(* Logix 5000 project; controller R400_500_XLS vendor 1 type 14 code 216 rev 31.11; software revision 31.01; part 5 of 32 *)
(* tags used below, declared in another part *)
   Abort1 : DINT;   // Not Used
   Cycles : UDT_CYCLE[11];
   CycleSequence : UDT_CYCLE_SEQUENCE;
   I_Pw_Tnk_Lvl_Sw_Deb : BOOL;   // Debounced pure water tank level switch (100ms)
   M : DINT[5];   // Memory Bits
   MinorFaultCheck : TIMER;
   MinorFaultRecord : FaultRecord;
   OneShot : DINT[1];
   ONS_FC01 : DINT;
   ONS_FC11 : DINT;
   ONS_FC12 : DINT;
   ONS_FC13 : DINT;
   ONS_FC64 : DINT;
   ONS_WSH30 : SINT;
   ONS_WSH35 : SINT;
   Service : DINT[2];   // Unused Service Mode Memory Bit
   String : STRING[50];   // String
   Tmr : TIMER[107];
   Unld_Door : DINT;
   BatteryLowWarning : BOOL;
   bFactoryResetCompleted : BOOL;
   bONSSerialModuleResetInhibit : BOOL;
   bONSSerialModuleSetInhibit : BOOL;
   bSerialModuleConfigureInhibit : BOOL;   // Configure if Serial Card is Inhibited or not
   Cfg_10_Modules : BOOL;   // Chassis is configured 10 slots
   Cfg_11_Modules : BOOL;
   Chassis_Size_Ret : DINT[3];
   Ctrlr_Status : DINT;
   Current_Screen : DINT;
   DateTime : DINT[7];
   DISABLE : BOOL;   // Disable bit
   EmailSMSInt : INT[8];   // Email & SMS Notification Integer
   EnDis_LabWasher : DINT;
   EnDis_LabWasher2 : DINT;
   Ethernet_Config_Msg : MESSAGE;
   F8 : REAL[6];
   I_Chem_Cond : DINT;   // Chemical water conductivity
   I_Chm_1_Lvl_Sw : BOOL;   // Chemical Pump #1 level switch
   I_Chm_2_Lvl_Sw : BOOL;   // Chemical Pump #2 level switch
   I_Chm_3_Lvl_Sw : BOOL;   // Chemical Pump #3 level switch
   I_Chm_4_Lvl_Sw : BOOL;   // Chemical Pump #4 level switch
   I_Dry_RTD : DINT;   // Drying RTD
   I_Final_Rinse_Cond : DINT;   // Final rinse water conductivity
   I_Ld_Dr_Cls_Sw : BOOL;   // Load door close
   I_Ld_Dr_Obs_Sw : BOOL;   // Load door obstruction switch
   I_MCR : BOOL;   // MCR input
   I_Mtr_Ovrld : BOOL;   // Motor overload
   I_Pump_Press : DINT;   // Recirculation pump pressure
   I_Pure_Water_Filling_Auth : BOOL;
   I_Pw_Tnk_Lvl_Sw : BOOL;   // Pure water tank level switch
   I_Pw_Tnk_RTD : DINT;   // Pure water tank RTD
   I_Pw_Tnk_Sft_Lvl_Sw : BOOL;   // Pure water tank safety level switch
   I_Shlf_Sw : BOOL;   // Shelf switch
   I_Smp_Lvl_Hgh : BOOL;   // Sump high level switch
   I_Smp_Lvl_Lw : BOOL;   // Sump low level switch
   I_Smp_RTD : DINT;   // Sump RTD
   I_Smp_Sft_Lvl_Sw : BOOL;   // Sump safety level switch
   I_Unld_Dr_Cls_Sw : BOOL;   // Unload door close
   I_Unld_Dr_Obs_Sw : BOOL;   // Unload door obstruction switch
   I_UnldDr_ClseSlnce_Bttn : BOOL;   // Door Close/ Silence button Unload Side
   I_UnldDr_Opn_Bttn : BOOL;   // Door Open button Unload side
   iSerialModuleActivateDeactivateInhibit : DINT;   // Set Bit 2 Of Word to Inhibited Serial M Reset Bit 2 Of Word to Un-inhibited
   L32E_ETH_Cfg : TIMER;   // Delay for Ethernet port initialization
   Language_English : STRING;
   MinorFaultBits : DINT;
   msg : BOOL[512];
   Msg_PwrUp : DINT;
   N13 : DINT;
   NOT_USED : SINT[3];
   ONS_WSH64 : SINT;
   previous_s108 : DINT;
   RD_CHASSIS_1 : MESSAGE;
   RD_CHASSIS_2 : MESSAGE;
   RemoteDisplayNumber : DINT;   // HMI connection
   sChangeLanguage : STRING;   // jplv09
   Screen_Ctrl : DINT;   // PLC Screen Request
   SimGenEnabled : BOOL;   // SimGen enable bit 1= Simgen ON
   Tpb : DINT[11];
   TpbImage : DINT[11];
   Unit : Hrdwre;   // Unit Configuration
   WR_CHASSIS_10 : MESSAGE;
   WR_CHASSIS_11 : MESSAGE;
(* MainProgram, continued *)

ROUTINE Inputs_10_Modules   (* ladder *)
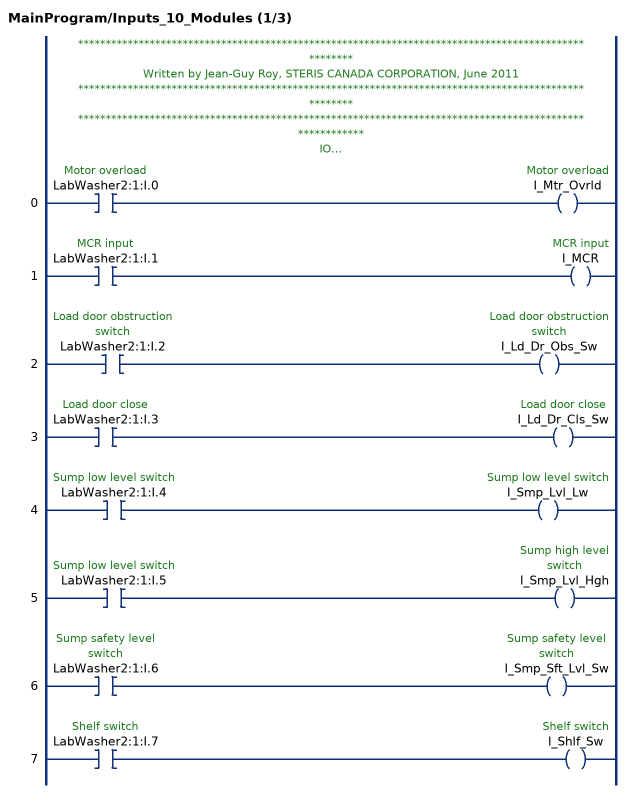
   // ****************************************************************************************************
   // Written by Jean-Guy Roy, STERIS CANADA CORPORATION, June 2011
   // ****************************************************************************************************
   // ********************************************************************************************************
   // IO1
   // ********************************************************************************************************
   0: XIC(LabWasher2:1:I.0)OTE(I_Mtr_Ovrld);
   1: XIC(LabWasher2:1:I.1)OTE(I_MCR);
   2: XIC(LabWasher2:1:I.2)OTE(I_Ld_Dr_Obs_Sw);
   3: XIC(LabWasher2:1:I.3)OTE(I_Ld_Dr_Cls_Sw);
   4: XIC(LabWasher2:1:I.4)OTE(I_Smp_Lvl_Lw);
   5: XIC(LabWasher2:1:I.5)OTE(I_Smp_Lvl_Hgh);
   6: XIC(LabWasher2:1:I.6)OTE(I_Smp_Sft_Lvl_Sw);
   7: XIC(LabWasher2:1:I.7)OTE(I_Shlf_Sw);
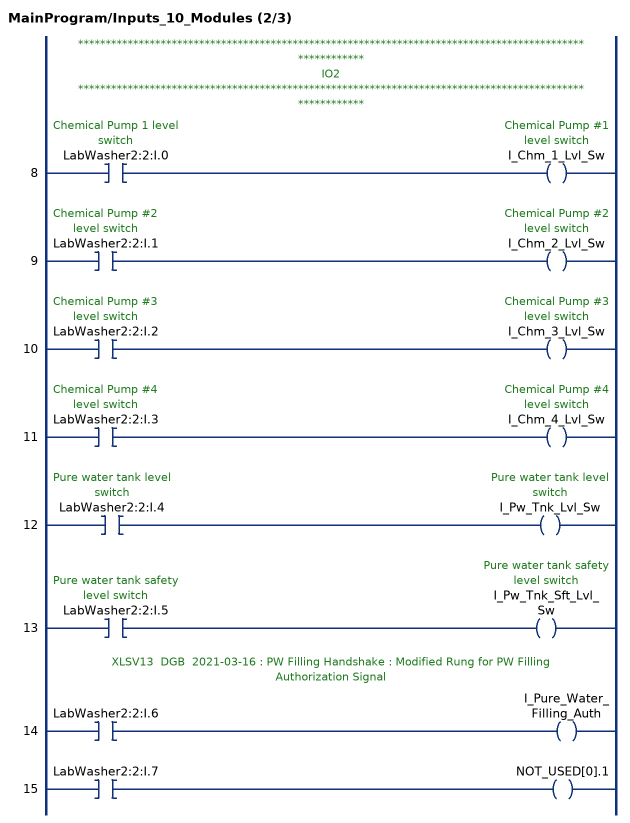
   // ********************************************************************************************************
   // IO2
   // ********************************************************************************************************
   8: XIC(LabWasher2:2:I.0)OTE(I_Chm_1_Lvl_Sw);
   9: XIC(LabWasher2:2:I.1)OTE(I_Chm_2_Lvl_Sw);
   10: XIC(LabWasher2:2:I.2)OTE(I_Chm_3_Lvl_Sw);
   11: XIC(LabWasher2:2:I.3)OTE(I_Chm_4_Lvl_Sw);
   12: XIC(LabWasher2:2:I.4)OTE(I_Pw_Tnk_Lvl_Sw);
   13: XIC(LabWasher2:2:I.5)OTE(I_Pw_Tnk_Sft_Lvl_Sw);
   // XLSV13  DGB  2021-03-16 : PW Filling Handshake : Modified Rung for PW Filling Authorization Signal
   14: XIC(LabWasher2:2:I.6)OTE(I_Pure_Water_Filling_Auth);
   15: XIC(LabWasher2:2:I.7)OTE(NOT_USED[0].1);
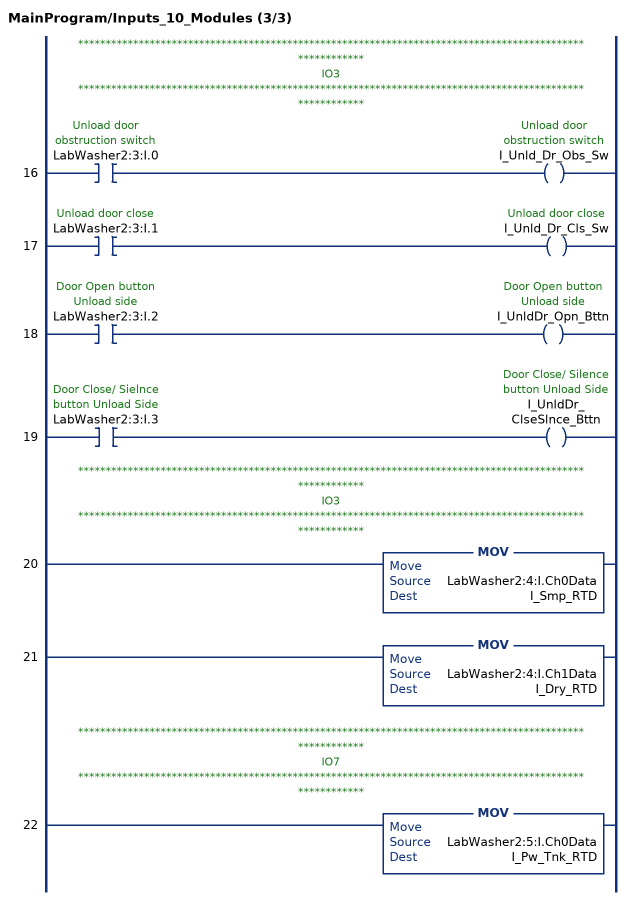
   // ********************************************************************************************************
   // IO3
   // ********************************************************************************************************
   16: XIC(LabWasher2:3:I.0)OTE(I_Unld_Dr_Obs_Sw);
   17: XIC(LabWasher2:3:I.1)OTE(I_Unld_Dr_Cls_Sw);
   18: XIC(LabWasher2:3:I.2)OTE(I_UnldDr_Opn_Bttn);
   19: XIC(LabWasher2:3:I.3)OTE(I_UnldDr_ClseSlnce_Bttn);
   // ********************************************************************************************************
   // IO3
   // ********************************************************************************************************
   20: MOV(LabWasher2:4:I.Ch0Data,I_Smp_RTD);
   21: MOV(LabWasher2:4:I.Ch1Data,I_Dry_RTD);
   // ********************************************************************************************************
   // IO7
   // ********************************************************************************************************
   22: MOV(LabWasher2:5:I.Ch0Data,I_Pw_Tnk_RTD);
END_ROUTINE

ROUTINE Inputs_Debounced   (* ladder *)
// This routine manages the debounced inputs
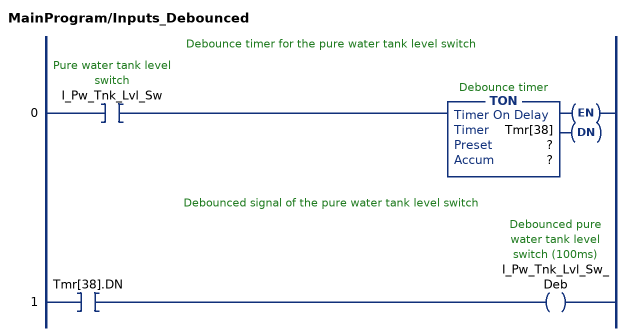
   // Debounce timer for the pure water tank level switch
   0: XIC(I_Pw_Tnk_Lvl_Sw)TON(Tmr[38],?,?);
   // Debounced signal of the pure water tank level switch
   1: XIC(Tmr[38].DN)OTE(I_Pw_Tnk_Lvl_Sw_Deb);
END_ROUTINE

ROUTINE Inputs_Smgn   (* ladder *)
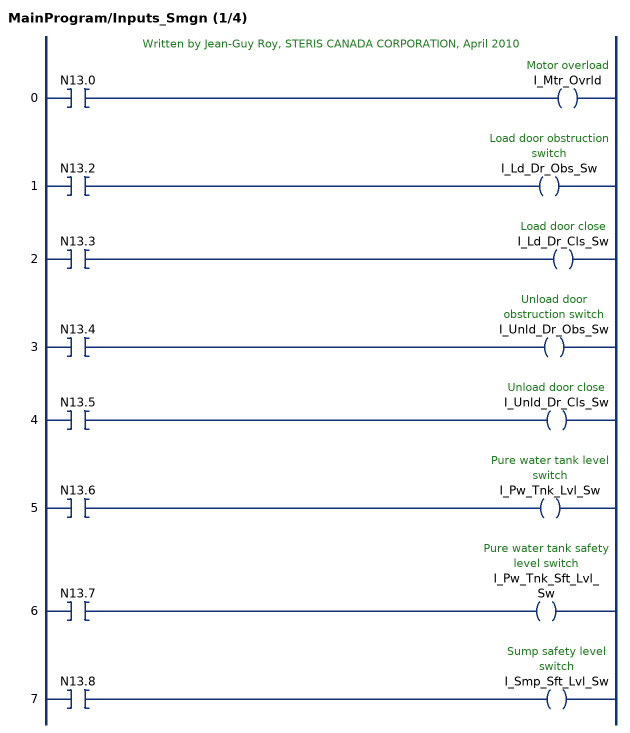
   // Written by Jean-Guy Roy, STERIS CANADA CORPORATION, April 2010
   0: XIC(N13.0)OTE(I_Mtr_Ovrld);
   1: XIC(N13.2)OTE(I_Ld_Dr_Obs_Sw);
   2: XIC(N13.3)OTE(I_Ld_Dr_Cls_Sw);
   3: XIC(N13.4)OTE(I_Unld_Dr_Obs_Sw);
   4: XIC(N13.5)OTE(I_Unld_Dr_Cls_Sw);
   5: XIC(N13.6)OTE(I_Pw_Tnk_Lvl_Sw);
   6: XIC(N13.7)OTE(I_Pw_Tnk_Sft_Lvl_Sw);
   7: XIC(N13.8)OTE(I_Smp_Sft_Lvl_Sw);
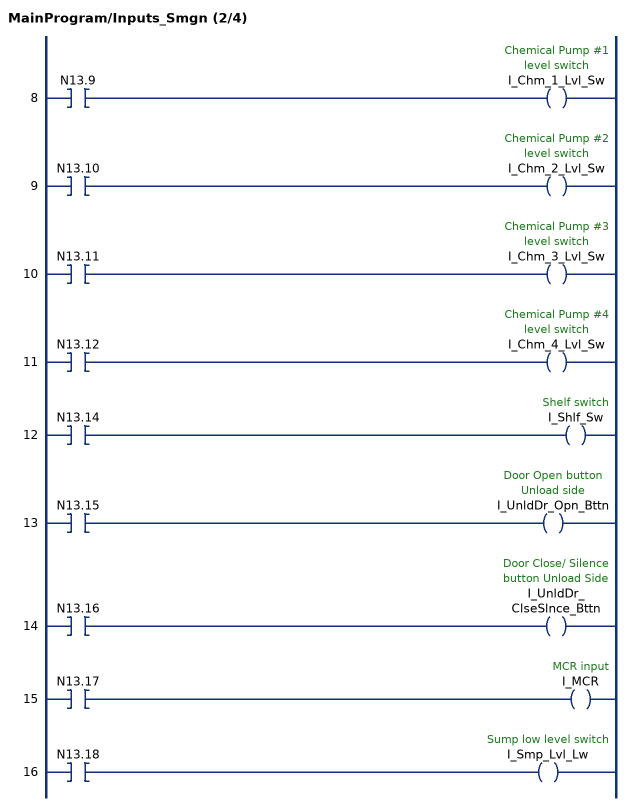
   8: XIC(N13.9)OTE(I_Chm_1_Lvl_Sw);
   9: XIC(N13.10)OTE(I_Chm_2_Lvl_Sw);
   10: XIC(N13.11)OTE(I_Chm_3_Lvl_Sw);
   11: XIC(N13.12)OTE(I_Chm_4_Lvl_Sw);
   12: XIC(N13.14)OTE(I_Shlf_Sw);
   13: XIC(N13.15)OTE(I_UnldDr_Opn_Bttn);
   14: XIC(N13.16)OTE(I_UnldDr_ClseSlnce_Bttn);
   15: XIC(N13.17)OTE(I_MCR);
   16: XIC(N13.18)OTE(I_Smp_Lvl_Lw);
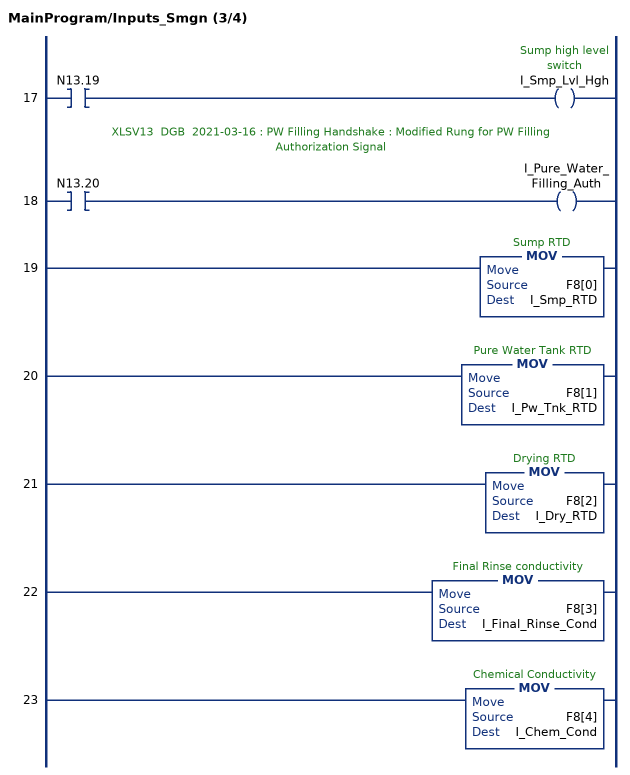
   17: XIC(N13.19)OTE(I_Smp_Lvl_Hgh);
   // XLSV13  DGB  2021-03-16 : PW Filling Handshake : Modified Rung for PW Filling Authorization Signal
   18: XIC(N13.20)OTE(I_Pure_Water_Filling_Auth);
   19: MOV(F8[0],I_Smp_RTD);
   20: MOV(F8[1],I_Pw_Tnk_RTD);
   21: MOV(F8[2],I_Dry_RTD);
   22: MOV(F8[3],I_Final_Rinse_Cond);
   23: MOV(F8[4],I_Chem_Cond);
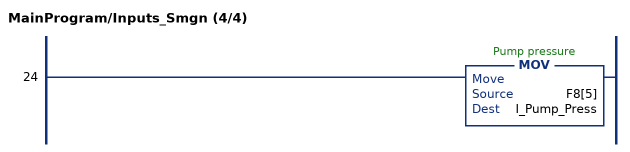
   24: MOV(F8[5],I_Pump_Press);
END_ROUTINE

ROUTINE MainRoutine   (* ladder *)
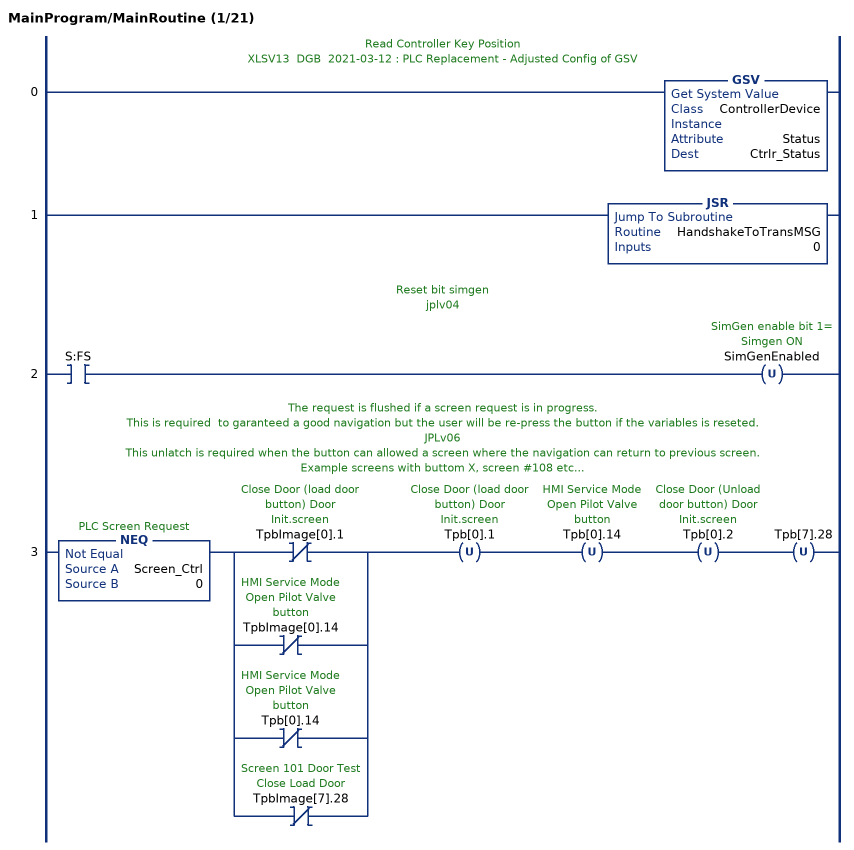
   // Read Controller Key Position
   // XLSV13  DGB  2021-03-12 : PLC Replacement - Adjusted Config of GSV
   0: GSV(ControllerDevice,,Status,Ctrlr_Status);
   1: JSR(HandshakeToTransMSG,0);
   // Reset bit simgen
   // jplv04
   2: XIC(S:FS)OTU(SimGenEnabled);
   // The request is flushed if a screen request is in progress.
   // This is required  to garanteed a good navigation but the user will be re-press the button if the variables is reseted.
   // JPLv06
   // This unlatch is required when the button can allowed a screen where the navigation can return to previous screen.
   // Example screens with buttom X, screen #108 etc...
   3: NEQ(Screen_Ctrl,0)[XIO(TpbImage[0].1) ,XIO(TpbImage[0].14) ,XIO(Tpb[0].14) ,XIO(TpbImage[7].28) ]OTU(Tpb[0].1)OTU(Tpb[0].14)OTU(Tpb[0].2)OTU(Tpb[7].28);
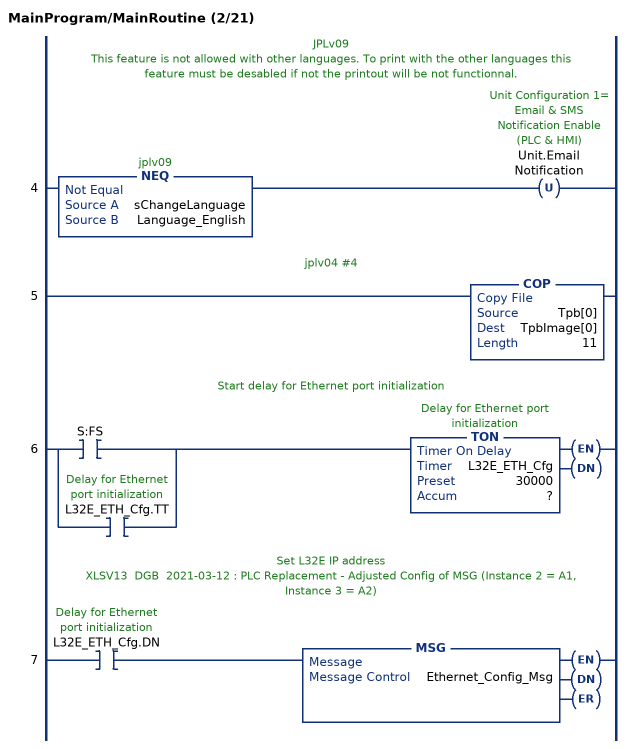
   // JPLv09
   // This feature is not allowed with other languages. To print with the other languages this feature must be desabled if not the printout will be not functionnal.
   4: NEQ(sChangeLanguage,Language_English)OTU(Unit.EmailNotification);
   // jplv04 #4
   5: COP(Tpb[0],TpbImage[0],11);
   // Start delay for Ethernet port initialization
   6: [XIC(S:FS) ,XIC(L32E_ETH_Cfg.TT) ]TON(L32E_ETH_Cfg,?,?);
   // Set L32E IP address
   // XLSV13  DGB  2021-03-12 : PLC Replacement - Adjusted Config of MSG (Instance 2 = A1, Instance 3 = A2)
   7: XIC(L32E_ETH_Cfg.DN)MSG(Ethernet_Config_Msg);
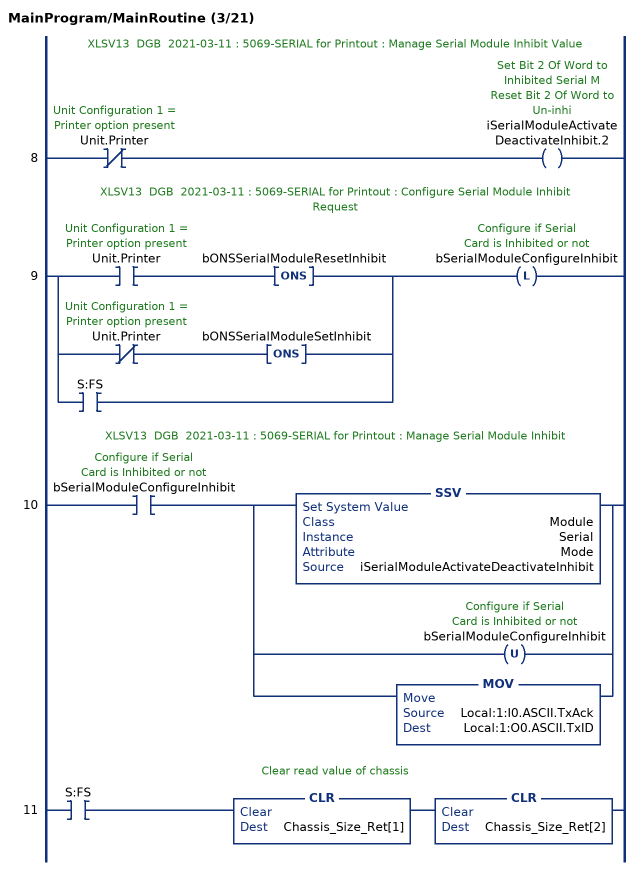
   // XLSV13  DGB  2021-03-11 : 5069-SERIAL for Printout : Manage Serial Module Inhibit Value
   8: XIO(Unit.Printer)OTE(iSerialModuleActivateDeactivateInhibit.2);
   // XLSV13  DGB  2021-03-11 : 5069-SERIAL for Printout : Configure Serial Module Inhibit Request
   9: [XIC(Unit.Printer) ONS(bONSSerialModuleResetInhibit) ,XIO(Unit.Printer) ONS(bONSSerialModuleSetInhibit) ,XIC(S:FS) ]OTL(bSerialModuleConfigureInhibit);
   // XLSV13  DGB  2021-03-11 : 5069-SERIAL for Printout : Manage Serial Module Inhibit
   10: XIC(bSerialModuleConfigureInhibit)[SSV(Module,Serial,Mode,iSerialModuleActivateDeactivateInhibit) ,OTU(bSerialModuleConfigureInhibit) ,MOV(Local:1:I0.ASCII.TxAck,Local:1:O0.ASCII.TxID) ];
   // Clear read value of chassis
   11: XIC(S:FS)CLR(Chassis_Size_Ret[1])CLR(Chassis_Size_Ret[2]);
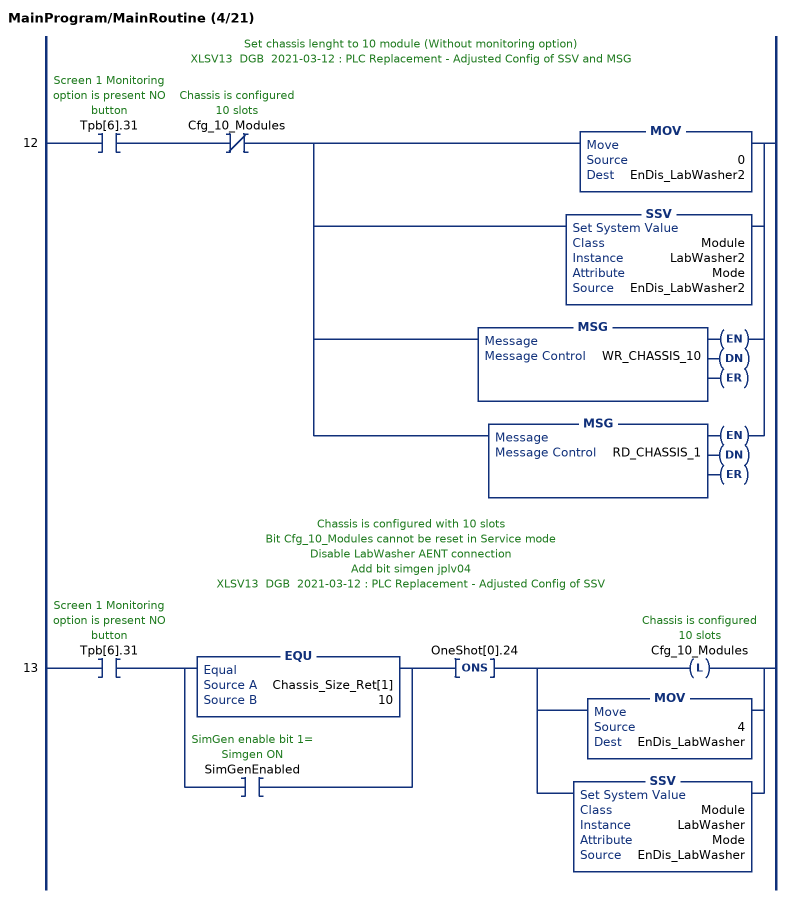
   // Set chassis lenght to 10 module (Without monitoring option)
   // XLSV13  DGB  2021-03-12 : PLC Replacement - Adjusted Config of SSV and MSG
   12: XIC(Tpb[6].31)XIO(Cfg_10_Modules)[MOV(0,EnDis_LabWasher2) ,SSV(Module,LabWasher2,Mode,EnDis_LabWasher2) ,MSG(WR_CHASSIS_10) ,MSG(RD_CHASSIS_1) ];
   // Chassis is configured with 10 slots
   // Bit Cfg_10_Modules cannot be reset in Service mode
   // Disable LabWasher AENT connection
   // Add bit simgen jplv04
   // XLSV13  DGB  2021-03-12 : PLC Replacement - Adjusted Config of SSV
   13: XIC(Tpb[6].31)[EQU(Chassis_Size_Ret[1],10) ,XIC(SimGenEnabled) ]ONS(OneShot[0].24)[OTL(Cfg_10_Modules) ,MOV(4,EnDis_LabWasher) ,SSV(Module,LabWasher,Mode,EnDis_LabWasher) ];
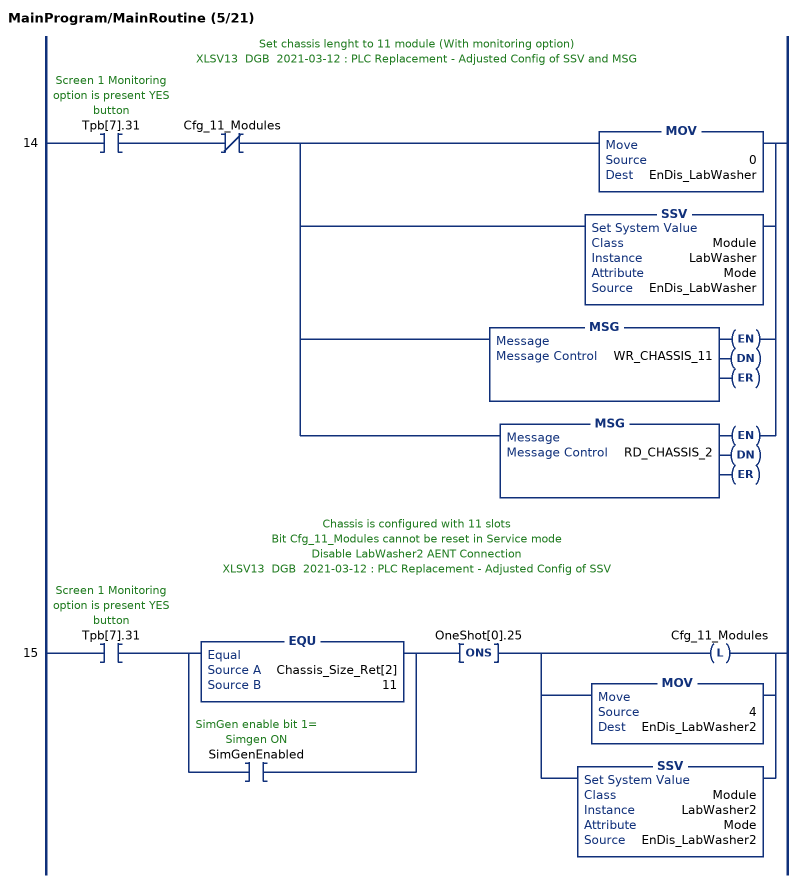
   // Set chassis lenght to 11 module (With monitoring option)
   // XLSV13  DGB  2021-03-12 : PLC Replacement - Adjusted Config of SSV and MSG
   14: XIC(Tpb[7].31)XIO(Cfg_11_Modules)[MOV(0,EnDis_LabWasher) ,SSV(Module,LabWasher,Mode,EnDis_LabWasher) ,MSG(WR_CHASSIS_11) ,MSG(RD_CHASSIS_2) ];
   // Chassis is configured with 11 slots
   // Bit Cfg_11_Modules cannot be reset in Service mode
   // Disable LabWasher2 AENT Connection
   // XLSV13  DGB  2021-03-12 : PLC Replacement - Adjusted Config of SSV
   15: XIC(Tpb[7].31)[EQU(Chassis_Size_Ret[2],11) ,XIC(SimGenEnabled) ]ONS(OneShot[0].25)[OTL(Cfg_11_Modules) ,MOV(4,EnDis_LabWasher2) ,SSV(Module,LabWasher2,Mode,EnDis_LabWasher2) ];
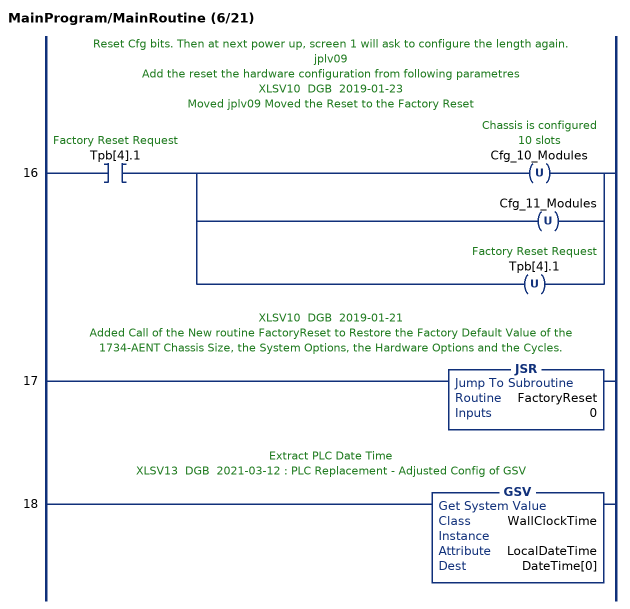
   // Reset Cfg bits. Then at next power up, screen 1 will ask to configure the length again.
   // jplv09
   // Add the reset the hardware configuration from following parametres
   // XLSV10  DGB  2019-01-23
   // Moved jplv09 Moved the Reset to the Factory Reset
   16: XIC(Tpb[4].1)[OTU(Cfg_10_Modules) ,OTU(Cfg_11_Modules) ,OTU(Tpb[4].1) ];
   // XLSV10  DGB  2019-01-21
   // Added Call of the New routine FactoryReset to Restore the Factory Default Value of the 1734-AENT Chassis Size, the System Options, the Hardware Options and the Cycles.
   17: JSR(FactoryReset,0);
   // Extract PLC Date Time
   // XLSV13  DGB  2021-03-12 : PLC Replacement - Adjusted Config of GSV
   18: GSV(WallClockTime,,LocalDateTime,DateTime[0]);
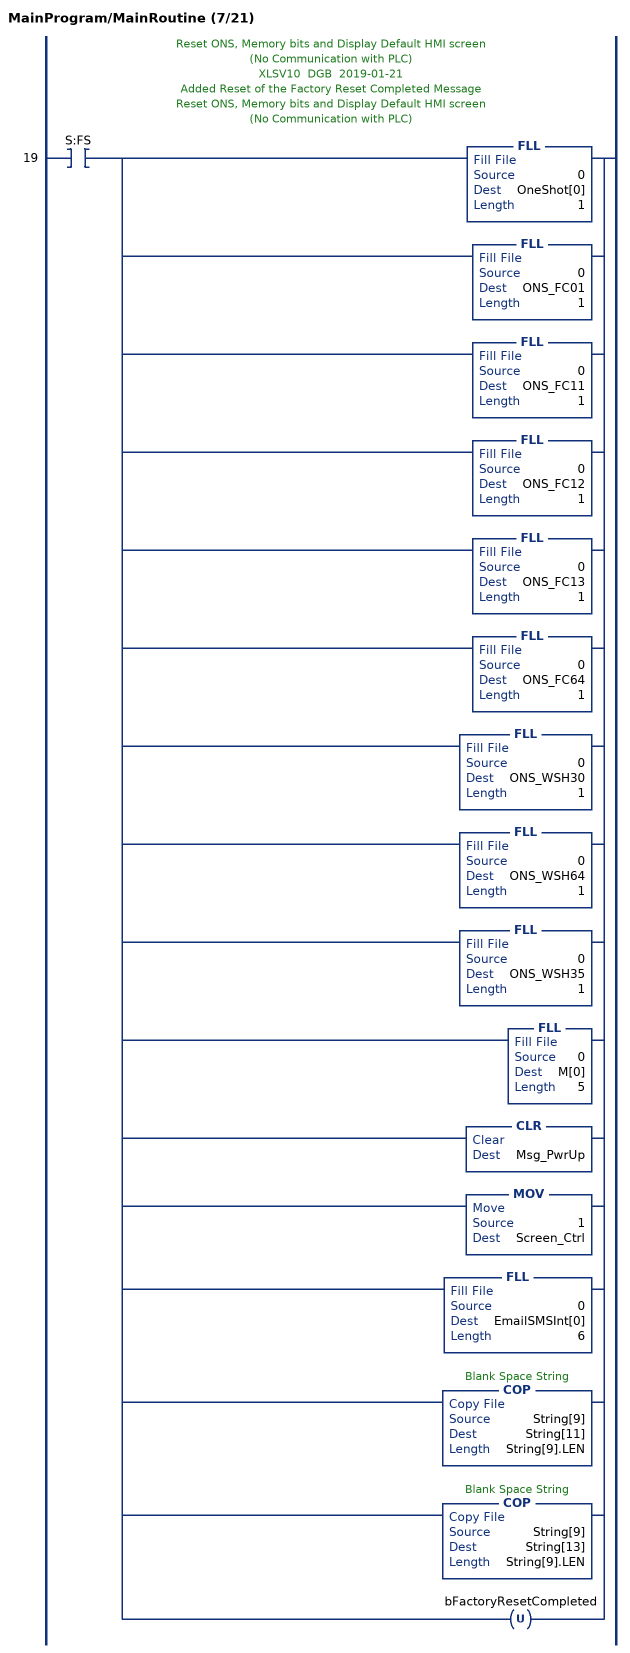
   // Reset ONS, Memory bits and Display Default HMI screen
   // (No Communication with PLC)
   // XLSV10  DGB  2019-01-21
   // Added Reset of the Factory Reset Completed Message
   // Reset ONS, Memory bits and Display Default HMI screen
   // (No Communication with PLC)
   19: XIC(S:FS)[FLL(0,OneShot[0],1) ,FLL(0,ONS_FC01,1) ,FLL(0,ONS_FC11,1) ,FLL(0,ONS_FC12,1) ,FLL(0,ONS_FC13,1) ,FLL(0,ONS_FC64,1) ,FLL(0,ONS_WSH30,1) ,FLL(0,ONS_WSH64,1) ,FLL(0,ONS_WSH35,1) ,FLL(0,M[0],5) ,CLR(Msg_PwrUp) ,MOV(1,Screen_Ctrl) ,FLL(0,EmailSMSInt[0],6) ,COP(String[9],String[11],String[9].LEN) ,COP(String[9],String[13],String[9].LEN) ,OTU(bFactoryResetCompleted) ];
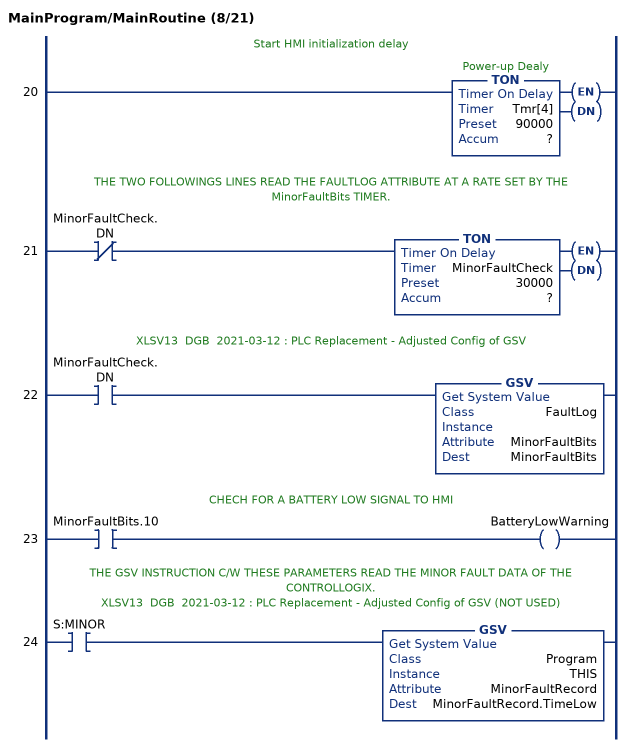
   // Start HMI initialization delay
   20: TON(Tmr[4],?,?);
   // THE TWO FOLLOWINGS LINES READ THE FAULTLOG ATTRIBUTE AT A RATE SET BY THE MinorFaultBits TIMER.
   21: XIO(MinorFaultCheck.DN)TON(MinorFaultCheck,?,?);
   // XLSV13  DGB  2021-03-12 : PLC Replacement - Adjusted Config of GSV
   22: XIC(MinorFaultCheck.DN)GSV(FaultLog,,MinorFaultBits,MinorFaultBits);
   // CHECH FOR A BATTERY LOW SIGNAL TO HMI
   23: XIC(MinorFaultBits.10)OTE(BatteryLowWarning);
   // THE GSV INSTRUCTION C/W THESE PARAMETERS READ THE MINOR FAULT DATA OF THE CONTROLLOGIX.
   // XLSV13  DGB  2021-03-12 : PLC Replacement - Adjusted Config of GSV (NOT USED)
   24: XIC(S:MINOR)GSV(Program,THIS,MinorFaultRecord,MinorFaultRecord.TimeLow);
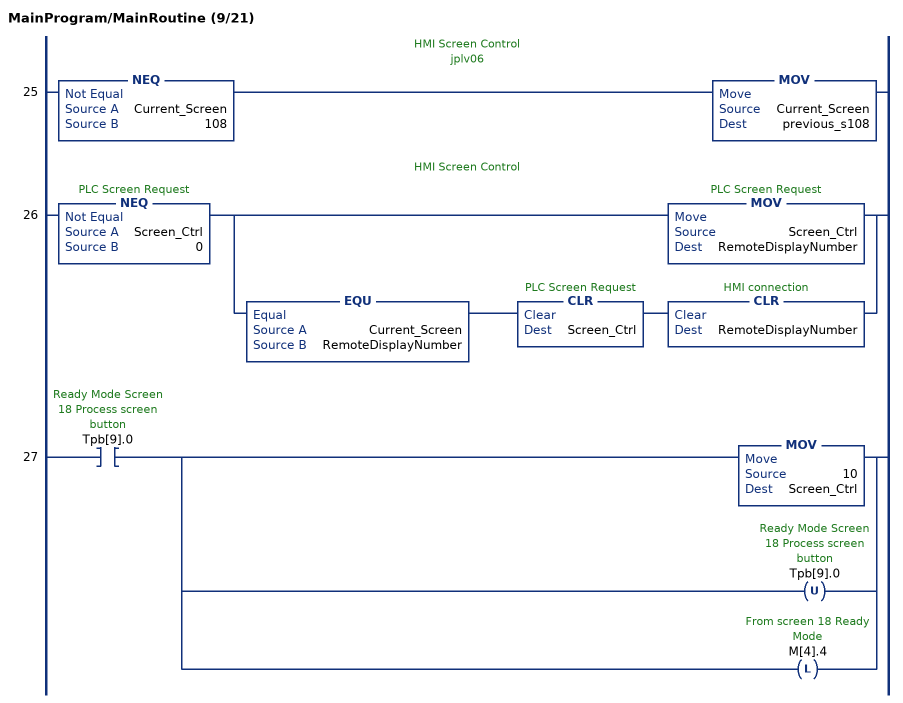
   // HMI Screen Control
   // jplv06
   25: NEQ(Current_Screen,108)MOV(Current_Screen,previous_s108);
   // HMI Screen Control
   26: NEQ(Screen_Ctrl,0)[MOV(Screen_Ctrl,RemoteDisplayNumber) ,EQU(Current_Screen,RemoteDisplayNumber) CLR(Screen_Ctrl) CLR(RemoteDisplayNumber) ];
   27: XIC(Tpb[9].0)[MOV(10,Screen_Ctrl) ,OTU(Tpb[9].0) ,OTL(M[4].4) ];
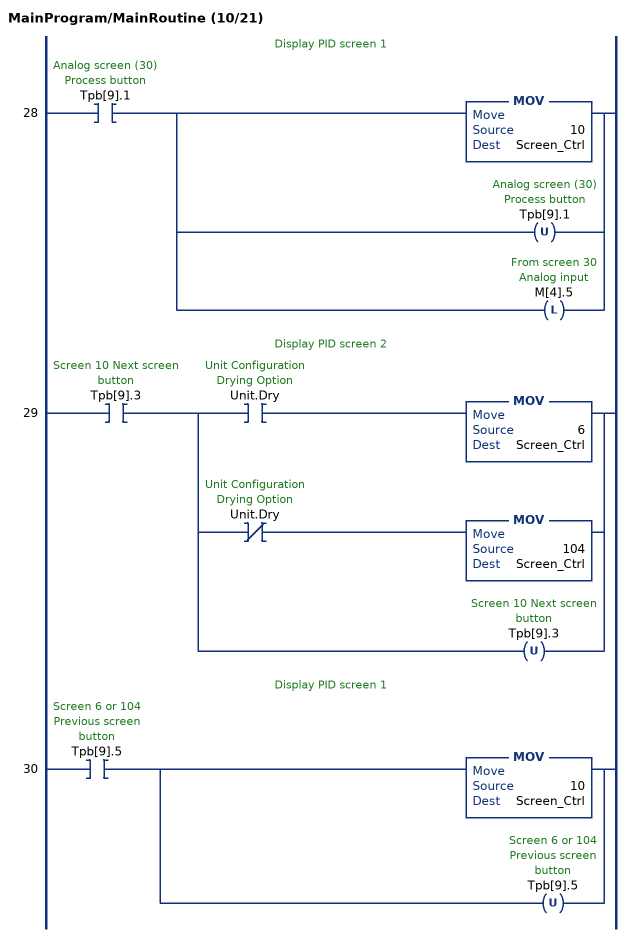
   // Display PID screen 1
   28: XIC(Tpb[9].1)[MOV(10,Screen_Ctrl) ,OTU(Tpb[9].1) ,OTL(M[4].5) ];
   // Display PID screen 2
   29: XIC(Tpb[9].3)[XIC(Unit.Dry) MOV(6,Screen_Ctrl) ,XIO(Unit.Dry) MOV(104,Screen_Ctrl) ,OTU(Tpb[9].3) ];
   // Display PID screen 1
   30: XIC(Tpb[9].5)[MOV(10,Screen_Ctrl) ,OTU(Tpb[9].5) ];
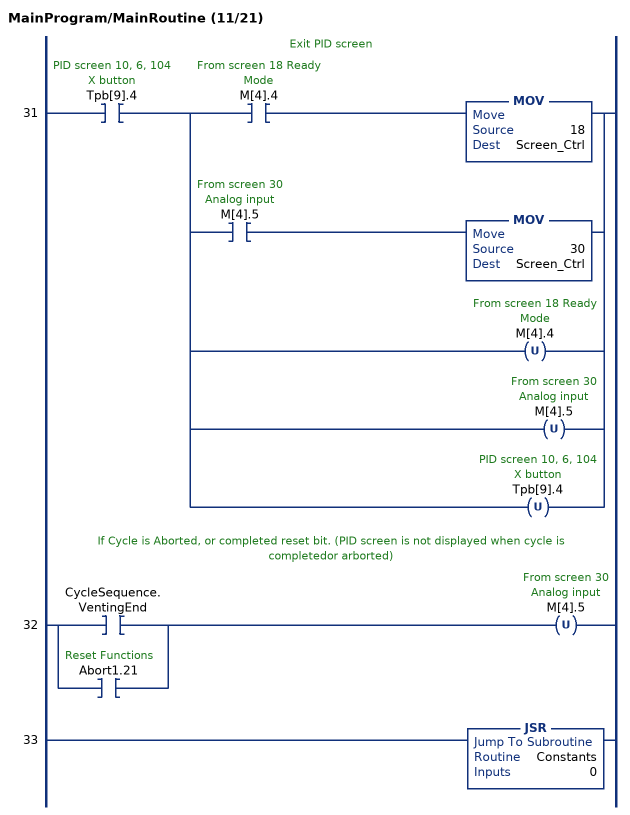
   // Exit PID screen
   31: XIC(Tpb[9].4)[XIC(M[4].4) MOV(18,Screen_Ctrl) ,XIC(M[4].5) MOV(30,Screen_Ctrl) ,OTU(M[4].4) ,OTU(M[4].5) ,OTU(Tpb[9].4) ];
   // If Cycle is Aborted, or completed reset bit. (PID screen is not displayed when cycle is completedor arborted)
   32: [XIC(CycleSequence.VentingEnd) ,XIC(Abort1.21) ]OTU(M[4].5);
   33: JSR(Constants,0);
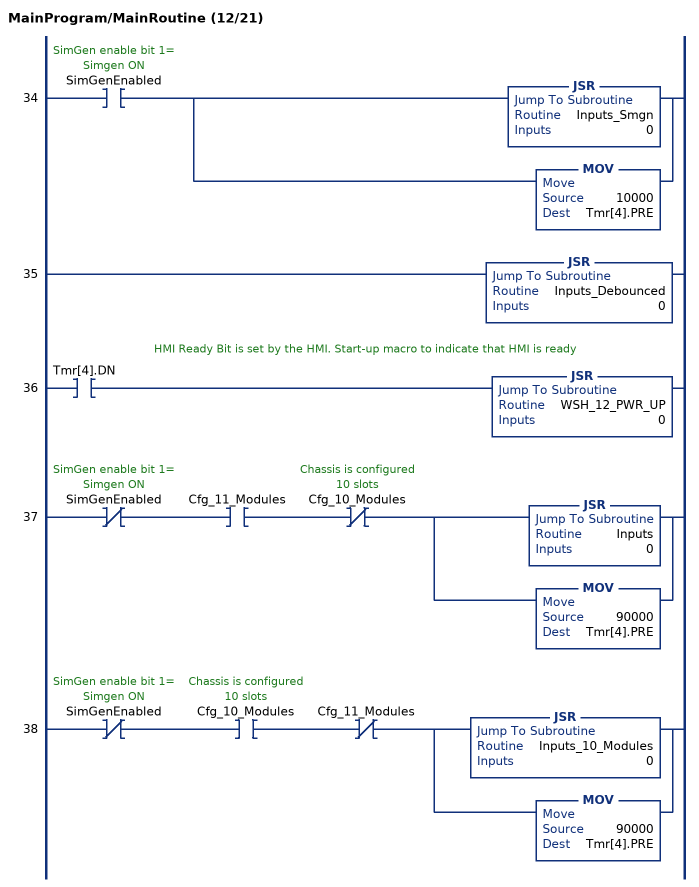
   34: XIC(SimGenEnabled)[JSR(Inputs_Smgn,0) ,MOV(10000,Tmr[4].PRE) ];
   35: JSR(Inputs_Debounced,0);
   // HMI Ready Bit is set by the HMI. Start-up macro to indicate that HMI is ready
   36: XIC(Tmr[4].DN)JSR(WSH_12_PWR_UP,0);
   37: XIO(SimGenEnabled)XIC(Cfg_11_Modules)XIO(Cfg_10_Modules)[JSR(Inputs,0) ,MOV(90000,Tmr[4].PRE) ];
   38: XIO(SimGenEnabled)XIC(Cfg_10_Modules)XIO(Cfg_11_Modules)[JSR(Inputs_10_Modules,0) ,MOV(90000,Tmr[4].PRE) ];
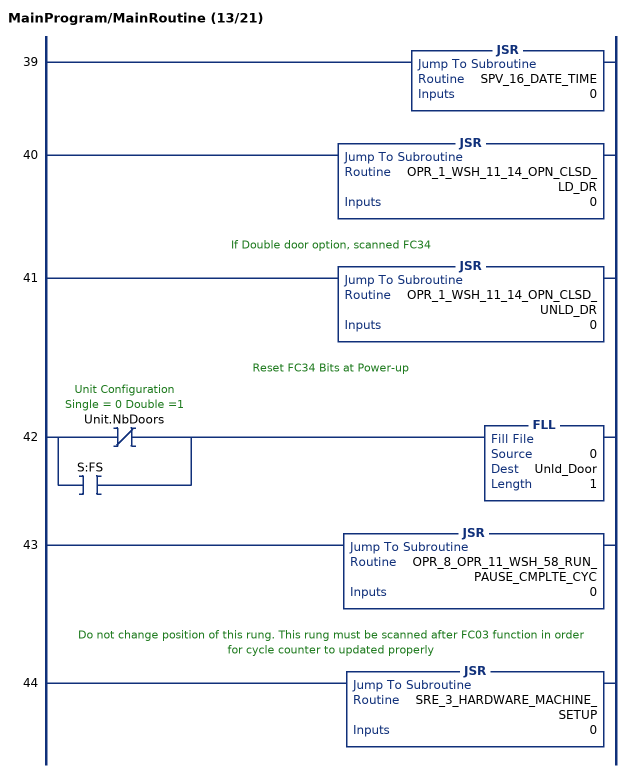
   39: JSR(SPV_16_DATE_TIME,0);
   40: JSR(OPR_1_WSH_11_14_OPN_CLSD_LD_DR,0);
   // If Double door option, scanned FC34
   41: JSR(OPR_1_WSH_11_14_OPN_CLSD_UNLD_DR,0);
   // Reset FC34 Bits at Power-up
   42: [XIO(Unit.NbDoors) ,XIC(S:FS) ]FLL(0,Unld_Door,1);
   43: JSR(OPR_8_OPR_11_WSH_58_RUN_PAUSE_CMPLTE_CYC,0);
   // Do not change position of this rung. This rung must be scanned after FC03 function in order for cycle counter to updated properly
   44: JSR(SRE_3_HARDWARE_MACHINE_SETUP,0);
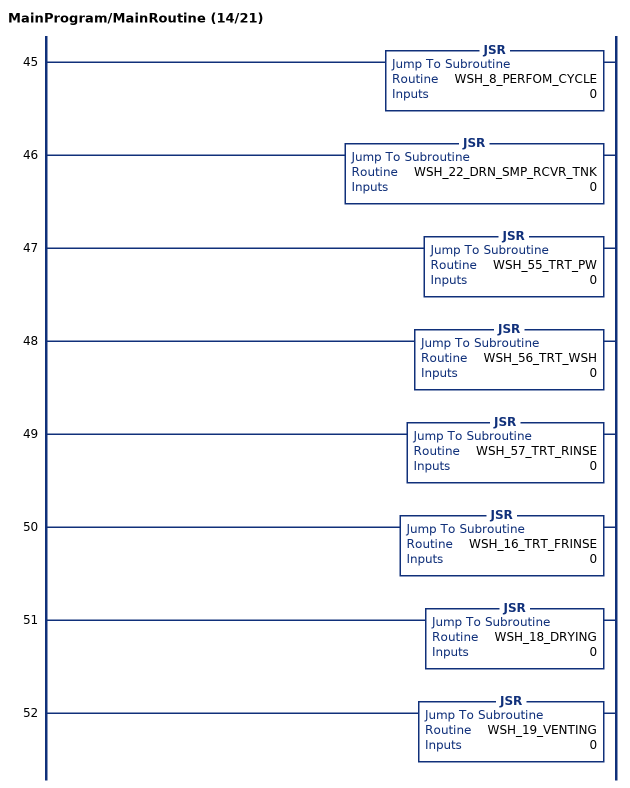
   45: JSR(WSH_8_PERFOM_CYCLE,0);
   46: JSR(WSH_22_DRN_SMP_RCVR_TNK,0);
   47: JSR(WSH_55_TRT_PW,0);
   48: JSR(WSH_56_TRT_WSH,0);
   49: JSR(WSH_57_TRT_RINSE,0);
   50: JSR(WSH_16_TRT_FRINSE,0);
   51: JSR(WSH_18_DRYING,0);
   52: JSR(WSH_19_VENTING,0);
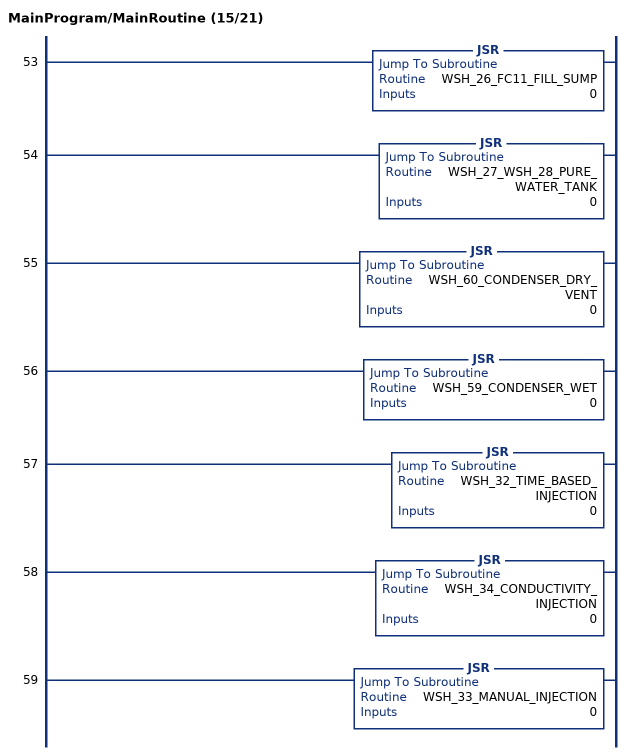
   53: JSR(WSH_26_FC11_FILL_SUMP,0);
   54: JSR(WSH_27_WSH_28_PURE_WATER_TANK,0);
   55: JSR(WSH_60_CONDENSER_DRY_VENT,0);
   56: JSR(WSH_59_CONDENSER_WET,0);
   57: JSR(WSH_32_TIME_BASED_INJECTION,0);
   58: JSR(WSH_34_CONDUCTIVITY_INJECTION,0);
   59: JSR(WSH_33_MANUAL_INJECTION,0);
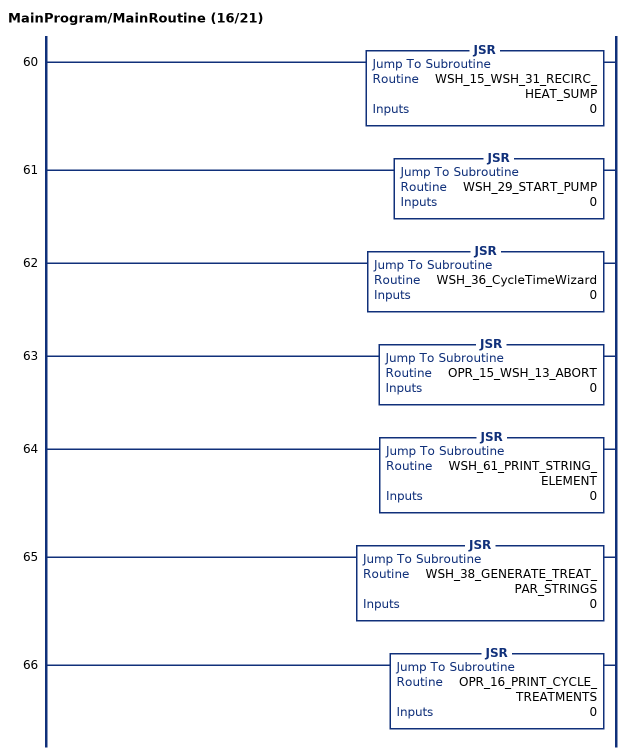
   60: JSR(WSH_15_WSH_31_RECIRC_HEAT_SUMP,0);
   61: JSR(WSH_29_START_PUMP,0);
   62: JSR(WSH_36_CycleTimeWizard,0);
   63: JSR(OPR_15_WSH_13_ABORT,0);
   64: JSR(WSH_61_PRINT_STRING_ELEMENT,0);
   65: JSR(WSH_38_GENERATE_TREAT_PAR_STRINGS,0);
   66: JSR(OPR_16_PRINT_CYCLE_TREATMENTS,0);
